// TIA Portal V20 export
Screen "180FX1Layout"  1276x673
  ScreenItem "Line_Header_X0_Y64" at 0,64 size 1276x0  Type=HmiLine
  ScreenItem "permanentareaborderrectangle" at 0,0 size 0x0  Type=HmiRectangle
  ScreenItem "Button_Back" at 2,2 size 90x60  Type=HmiButton
  ScreenItem "Move_Legend" at 1182,2 size 90x60  Type=HmiButton
  ScreenItem "Fusszeile_Button_ManualOPMode1_2" at 279,2 size 90x60  Type=HmiButton
  ScreenItem "文本域_3" at 1107,71 size 139x22  Type=HmiTextBox
  ScreenItem "文本域_1" at 1107,160 size 156x23  Type=HmiTextBox
  ScreenItem "文本域_22" at 1124,283 size 104x23  Type=HmiTextBox
  ScreenItem "面板容器_2" at 1090,4 size 88x58  Type=HmiFaceplateContainer
  ScreenItem "OPMode1_Blocked" at 1164,6 size 14x14  Type=HmiGraphicView
  ScreenItem "OPMode4_Foreground_Blocked" at 1090,5 size 88x58  Type=HmiGraphicView
  ScreenItem "Fusszeile_Button_ManualOPMode1_1" at 95,2 size 90x60  Type=HmiButton
  ScreenItem "Graphic view_1" at 119,217 size 756x259  Type=HmiGraphicView
  ScreenItem "Line_2" at 174,159 size 40x96  Type=HmiLine
  ScreenItem "Line_6" at 799,329 size 128x0  Type=HmiLine
  ScreenItem "Fusszeile_Button_ManualOPMode1_3" at 187,2 size 90x60  Type=HmiButton
  ScreenItem "文本域_6" at 144,91 size 140x40  Type=HmiTextBox
  ScreenItem "文本域_12" at 929,305 size 100x40  Type=HmiTextBox
  ScreenItem "文本域_13" at 514,91 size 140x20  Type=HmiTextBox
  ScreenItem "文本域_14" at 936,-172 size 140x40  Type=HmiTextBox
  ScreenItem "文本域_15" at 914,173 size 140x40  Type=HmiTextBox
  ScreenItem "Title_ScreenOverview_X390_Y2_1" at 384,5 size 510x57  Type=HmiTextBox
  ScreenItem "Line_12" at 831,210 size 82x77  Type=HmiLine
  ScreenItem "文本域_24" at 685,91 size 140x20  Type=HmiTextBox
  ScreenItem "文本域_26" at 914,418 size 140x40  Type=HmiTextBox
  ScreenItem "Line_14" at 745,139 size 43x179  Type=HmiLine
  ScreenItem "Line_15" at 741,342 size 47x197  Type=HmiLine
  ScreenItem "Line_19" at 830,372 size 82x54  Type=HmiLine
  ScreenItem "Line_1" at 585,338 size 103x201  Type=HmiLine
  ScreenItem "Line_3" at 574,136 size 97x122  Type=HmiLine
  ScreenItem "面板容器_5" at 144,133 size 143x50  Type=HmiFaceplateContainer
  ScreenItem "面板容器_10" at 514,111 size 153x58  Type=HmiFaceplateContainer
  ScreenItem "面板容器_15" at 914,458 size 149x54  Type=HmiFaceplateContainer
  ScreenItem "面板容器_6" at 914,215 size 149x54  Type=HmiFaceplateContainer
  ScreenItem "Faceplate container_6" at 949,346 size 59x45  Type=HmiFaceplateContainer
  ScreenItem "面板容器_4" at 685,112 size 142x51  Type=HmiFaceplateContainer
  ScreenItem "面板容器_1" at 685,559 size 142x51  Type=HmiFaceplateContainer
  ScreenItem "Faceplate container_7" at 554,579 size 59x45  Type=HmiFaceplateContainer
  ScreenItem "面板容器_23" at 1178,251 size 96x32  Type=HmiFaceplateContainer
  ScreenItem "面板容器_22" at 1068,251 size 96x32  Type=HmiFaceplateContainer
  ScreenItem "LSicar_Valve8Pos_LeftHomeRightWork_WithPB_5" at 1099,95 size 160x53  Type=HmiFaceplateContainer
  ScreenItem "LSicar_Valve8Pos_LeftHomeRightWork_WithPB_1" at 1099,183 size 160x53  Type=HmiFaceplateContainer
  ScreenItem "文本域_20" at 875,91 size 140x20  Type=HmiTextBox
  ScreenItem "文本域_11" at 875,539 size 140x20  Type=HmiTextBox
  ScreenItem "面板容器_9" at 875,559 size 148x58  Type=HmiFaceplateContainer
  ScreenItem "Line_4" at 813,400 size 69x137  Type=HmiLine
  ScreenItem "Line_5" at 817,120 size 71x139  Type=HmiLine
  ScreenItem "Line_Header_X0_Y64_1" at 0,64 size 1276x0  Type=HmiLine
  ScreenItem "文本域_27" at -1,126 size 120x40  Type=HmiTextBox
  ScreenItem "文本域_5" at -1,82 size 120x40  Type=HmiTextBox
  ScreenItem "文本域_25" at 685,539 size 140x20  Type=HmiTextBox
  ScreenItem "文本域_8" at 534,539 size 100x40  Type=HmiTextBox
  ScreenItem "面板容器_7" at 875,111 size 148x58  Type=HmiFaceplateContainer
